(* IEC 61131-3 sources: llm-plc-st-eval/data/calibracion/claude-sonnet-4-6/B1/zero_shot, 3 files *)

(* ---- ejec_1.st ---- *)
```pascal
FUNCTION_BLOCK FB_Motor
VAR_INPUT
    btnMarcha : BOOL; (* Botón de marcha: TRUE = pulsado *)
    btnParo   : BOOL; (* Botón de paro: TRUE = pulsado *)
    btnEmerg  : BOOL; (* Paro de emergencia: TRUE = activado *)
END_VAR

VAR_OUTPUT
    motorOn : BOOL; (* Salida al contactor del motor *)
END_VAR

VAR
    bloqueEmerg : BOOL; (* Enclavamiento por emergencia *)
END_VAR

(*
    Lógica de control:
    1. Si se activa la emergencia → parar motor y bloquear rearranque.
    2. El bloqueo de emergencia solo se libera cuando btnEmerg vuelve
       a FALSE (emergencia restablecida) Y el botón de marcha NO está
       pulsado, evitando un arranque automático no deseado.
    3. Paro normal: btnParo detiene el motor sin bloquear el rearranque.
    4. Arranque: btnMarcha activa el motor si no hay bloqueo ni paro.
    5. Auto-retención: motorOn se mantiene mediante su propio estado.
*)

(* --- Gestión del enclavamiento de emergencia --- *)
IF btnEmerg THEN
    (* Activar bloqueo al detectar emergencia *)
    bloqueEmerg := TRUE;
ELSIF NOT btnEmerg AND NOT btnMarcha THEN
    (* Liberar bloqueo solo cuando la emergencia se restablece
       y el botón de marcha no está presionado *)
    bloqueEmerg := FALSE;
END_IF;

(* --- Lógica de arranque / paro del motor --- *)
IF btnEmerg OR btnParo OR bloqueEmerg THEN
    (* Prioridad de paro: emergencia, paro normal o bloqueo activo *)
    motorOn := FALSE;
ELSIF btnMarcha AND NOT bloqueEmerg THEN
    (* Arranque: condición de marcha sin bloqueo *)
    motorOn := TRUE;
END_IF;
(* Auto-retención implícita: motorOn conserva su valor TRUE
   mientras no se active ninguna condición de paro *)

END_FUNCTION_BLOCK
```

(* ---- ejec_2.st ---- *)
```pascal
FUNCTION_BLOCK FB_Motor
VAR_INPUT
    btnMarcha : BOOL; (* Botón de marcha: TRUE = pulsado *)
    btnParo   : BOOL; (* Botón de paro: TRUE = pulsado   *)
    btnEmerg  : BOOL; (* Paro de emergencia: TRUE = activo *)
END_VAR

VAR_OUTPUT
    motorOn : BOOL; (* TRUE = motor en marcha *)
END_VAR

VAR
    bloqueado : BOOL; (* Enclavamiento post-emergencia *)
END_VAR

(*
    Lógica de control:
    1. Si se activa la emergencia: parar motor y activar enclavamiento.
    2. Si el enclavamiento está activo: el motor no puede arrancar.
       El enclavamiento solo se libera cuando btnEmerg vuelve a FALSE
       Y btnMarcha NO está pulsado (evita rearranque automático).
    3. Si se pulsa paro: apagar motor (sin enclavamiento).
    4. Si se pulsa marcha y no hay enclavamiento ni paro: arrancar y
       mantener motor (auto-retención por lógica de estado).
*)

(* --- Paso 1: Gestión de emergencia --- *)
IF btnEmerg THEN
    motorOn   := FALSE;
    bloqueado := TRUE;  (* Activar enclavamiento *)
END_IF;

(* --- Paso 2: Liberación del enclavamiento ---
   Solo se libera cuando la emergencia se ha retirado
   Y el botón de marcha no está pulsado en ese instante *)
IF bloqueado AND NOT btnEmerg AND NOT btnMarcha THEN
    bloqueado := FALSE;
END_IF;

(* --- Paso 3 y 4: Control normal (solo si no hay emergencia activa
   ni enclavamiento vigente) --- *)
IF NOT btnEmerg AND NOT bloqueado THEN

    IF btnParo THEN
        (* Paro normal: apagar motor *)
        motorOn := FALSE;

    ELSIF btnMarcha THEN
        (* Arranque: encender motor *)
        motorOn := TRUE;

    (* Si ningún botón está pulsado, motorOn conserva su estado
       anterior (auto-retención implícita por variable de estado) *)
    END_IF;

END_IF;
```

(* ---- ejec_3.st ---- *)
```pascal
FUNCTION_BLOCK FB_Motor
VAR_INPUT
    btnMarcha : BOOL; (* Botón de marcha: TRUE = pulsado *)
    btnParo   : BOOL; (* Botón de paro: TRUE = pulsado *)
    btnEmerg  : BOOL; (* Paro de emergencia: TRUE = activado *)
END_VAR

VAR_OUTPUT
    motorOn : BOOL; (* Salida al contactor del motor *)
END_VAR

VAR
    bloqueEmerg : BOOL := FALSE; (* Bloqueo activo tras emergencia *)
END_VAR

(*
    Lógica de control:
    1. Si se activa la emergencia → parar motor y activar bloqueo.
    2. El bloqueo se libera SOLO cuando btnEmerg vuelve a FALSE
       Y btnMarcha NO está pulsado (evita rearranque automático).
    3. Paro normal → apagar motor (sin bloqueo).
    4. Marcha → encender motor si no hay bloqueo ni paro activo.
    5. Autoenclavamiento: motorOn se mantiene al soltar btnMarcha.
*)

(* --- Paso 1: Gestión del bloqueo por emergencia --- *)
IF btnEmerg THEN
    (* Emergencia activa: bloquear y apagar *)
    bloqueEmerg := TRUE;
    motorOn     := FALSE;

ELSIF bloqueEmerg THEN
    (* Emergencia retirada: liberar bloqueo solo si btnMarcha no está pulsado *)
    IF NOT btnMarcha THEN
        bloqueEmerg := FALSE;
    END_IF;
    (* Motor permanece apagado mientras dure el bloqueo *)
    motorOn := FALSE;

ELSE
    (* --- Paso 2: Operación normal (sin emergencia ni bloqueo) --- *)

    IF btnParo THEN
        (* Paro normal: apagar motor *)
        motorOn := FALSE;

    ELSIF btnMarcha THEN
        (* Marcha: encender motor *)
        motorOn := TRUE;

    END_IF;
    (* Si ningún botón está pulsado, motorOn conserva su valor → autoenclavamiento *)

END_IF;
```
